(* IEC 61131-3 sources: kns-pump-station/tests/POUs/Field/FB_PlcStartAdoption_Test, 4 files *)

(* ---- FB_PlcStartAdoption_Test.decl.st ---- *)
// Назначение: набор coUnit — подхват работающего насоса при старте ПЛК в порядке вызова сгенерированного
//             PRG_Devices: ES301 (link_power) вызывается раньше насосов, его значение в первом вызове берётся
//             без задержки DI (plc-process-lib, DI-1), поэтому первый вызов FB_MotorVfd видит напряжение и
//             подхватывает работающий по ОС насос с запросом станции. Обратный порядок (как по dev_no в
//             iolistgen 0.1.0) показывает, зачем порядок нужен: без напряжения подхват кончается остановом.
//             Устройства — настоящие ФБ библиотеки с параметрами проекта (GVL_CfgProject).
// Автор:      kr0nsch
// Версия:     0.1.0
// Документ:   docs/DESIGN.md, разделы 4.6, 7; docs/04_algorithms.md, раздел 13.3; docs/ASSUMPTIONS.md, И3
FUNCTION_BLOCK FB_PlcStartAdoption_Test EXTENDS coUnit.FB_TestSuite
VAR CONSTANT
    R_SPEED_PCT : REAL := 70.0;     // частота работающего ПЧ, %
END_VAR

(* ---- AdoptedInGeneratedOrder.method.decl.st ---- *)
// Сгенерированный порядок (ES301, затем P101): насос работает по ОС (реле «Работа» ПЧ, xFbFromComm = FALSE),
// станция подхватила его запросом (xAutoRun из GVL_IO.xP101_RFB в первом цикле) — первый вызов P101 видит
// напряжение, насос в Running с командой xQRun, пуск не засчитан; через 5 с — так же, без отказов
METHOD PRIVATE AdoptedInGeneratedOrder
VAR
    fbTime   : PL.FB_FakeTime;          // подменное время, старт 1 ч
    stDiCmd  : PL.ST_DigitalInputCmd;   // GVL_Hmi.stES301Cmd
    stDiCfg  : PL.ST_DigitalInputCfg;   // GVL_Persist.stES301Cfg
    stMotCmd : PL.ST_MotorCmd;          // GVL_Hmi.stP101Cmd
    stMotCfg : PL.ST_MotorCfg;          // GVL_Persist.stP101Cfg
    stMotRet : PL.ST_DeviceRetain;      // GVL_Persist.stP101Retain
    uiStep   : UINT;                    // шаг
END_VAR
VAR_INST
    fbES301  : PL.FB_DigitalInput;      // GVL_Devices.fbES301
    fbP101   : PL.FB_MotorVfd;          // GVL_Devices.fbP101
END_VAR

(* ---- AdoptedInGeneratedOrder.method.impl.st ---- *)
coUnit.TEST('PlcStartAdoption_AdoptedInGeneratedOrder_A13');

stDiCfg := GVL_CfgProject.stES301Cfg;
stMotCfg := GVL_CfgProject.stP101Cfg;
stMotRet.eRemoteMode := PL.E_DeviceMode.Auto;
// первый вызов (старт ПЛК) в порядке PRG_Devices: ES301, затем P101 с напряжением от ES301
fbTime.Advance(tStep := T#100MS);
fbES301(xIn := TRUE, xChannelFault := FALSE, itfTime := fbTime, stCmd := stDiCmd, stCfg := stDiCfg);
fbP101(xAutoRun := TRUE, rSpeedSpAuto_pct := R_SPEED_PCT, xFbRun := TRUE, xExtFault := FALSE, xLocal := FALSE,
       xPowerOk := fbES301.xValue, xCommOk := TRUE, xVfdRunning := TRUE, xVfdReady := TRUE, xVfdFault := FALSE,
       rSpeedAct_pct := R_SPEED_PCT, itfTime := fbTime, stCmd := stMotCmd, stCfg := stMotCfg, stRetain := stMotRet);
AssertTrue(Condition := fbES301.xValue, Message := 'first call: power value without DI delay');
AssertTrue(Condition := fbP101.stSts.eState = PL.E_MotorState.Running, Message := 'first call: adopted');
AssertTrue(Condition := fbP101.xQRun, Message := 'first call: run command kept');

// дальше — 5 с по 100 мс в том же порядке
FOR uiStep := 1 TO 50 DO
    fbTime.Advance(tStep := T#100MS);
    fbES301(xIn := TRUE, xChannelFault := FALSE, itfTime := fbTime, stCmd := stDiCmd, stCfg := stDiCfg);
    fbP101(xAutoRun := TRUE, rSpeedSpAuto_pct := R_SPEED_PCT, xFbRun := TRUE, xExtFault := FALSE, xLocal := FALSE,
           xPowerOk := fbES301.xValue, xCommOk := TRUE, xVfdRunning := TRUE, xVfdReady := TRUE, xVfdFault := FALSE,
           rSpeedAct_pct := R_SPEED_PCT, itfTime := fbTime, stCmd := stMotCmd, stCfg := stMotCfg,
           stRetain := stMotRet);
END_FOR
AssertTrue(Condition := fbP101.stSts.eState = PL.E_MotorState.Running, Message := 'after 5 s: still running');
AssertTrue(Condition := fbP101.xQRun, Message := 'after 5 s: run command kept');
AssertEquals_UDINT(Expected := 0, Actual := stMotRet.udiOpCount, Message := 'adoption is not a start');
AssertEquals_WORD(Expected := 0, Actual := fbP101.stSts.stCommon.wFault, Message := 'no fault');

coUnit.TEST_FINISHED();

(* ---- PowerDeviceAfterPumpStopsRunningPump.method.decl.st ---- *)
// Обратный порядок (P101 раньше ES301, как по dev_no без учёта link_power): в первом вызове P101 значение
// ES301 ещё не посчитано (FALSE) — подхват сразу сменяется остановом «нет напряжения», команда снята.
// Поэтому порядок вызова — свойство сгенерированного PRG_Devices (проверяет и test_generate.py)
METHOD PRIVATE PowerDeviceAfterPumpStopsRunningPump
VAR
    fbTime   : PL.FB_FakeTime;          // подменное время, старт 1 ч
    stDiCmd  : PL.ST_DigitalInputCmd;   // GVL_Hmi.stES301Cmd
    stDiCfg  : PL.ST_DigitalInputCfg;   // GVL_Persist.stES301Cfg
    stMotCmd : PL.ST_MotorCmd;          // GVL_Hmi.stP101Cmd
    stMotCfg : PL.ST_MotorCfg;          // GVL_Persist.stP101Cfg
    stMotRet : PL.ST_DeviceRetain;      // GVL_Persist.stP101Retain
END_VAR
VAR_INST
    fbES301  : PL.FB_DigitalInput;      // GVL_Devices.fbES301
    fbP101   : PL.FB_MotorVfd;          // GVL_Devices.fbP101
END_VAR
